(* CODESYS project JobManager.xml

Project tree, tasks and I/O mapping:
  visualisation JobManager
*)

// /JobManager
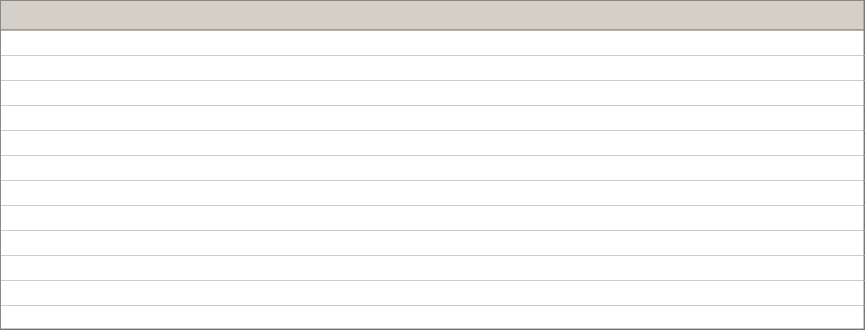
VISUALIZATION JobManager  // 865x330
    Table (0,0 865x330), data array: PRG_VisuTask_10ms._fbJobMgrCtrl._ascJobs
        p1128707560: cMaxNbrOfJobs
        p1014161805: GVL_Constant.cMaxNbrOfJobs - 1 + 1
        p3854506369: PRG_VisuTask_10ms._fbJobMgrCtrl._ascJobs[INDEX].eJobType
        p1892666644: PRG_VisuTask_10ms._fbJobMgrCtrl._ascJobs[INDEX].eJobState
        p338671338: PRG_VisuTask_10ms._fbJobMgrCtrl._ascJobs[INDEX].eJobPriority
        p2170511999: PRG_VisuTask_10ms._fbJobMgrCtrl._ascJobs[INDEX].eFrame
        p3723444502: PRG_VisuTask_10ms._fbJobMgrCtrl._ascJobs[INDEX].eSide
        p2232123230: Job Type
        p511219082: Job State
        p1755163831: Job Priority
        p4092479075: UserFrame
END_VISUALIZATION
